// TIA Portal V21 export
// export: Created 2026-11-10T07:35:10.4726746Z, ExportSetting WithDefaults, DisplayName Totally Integrated Automation Portal, DisplayVersion V21 Update 3, DisplayName STEP 7 Professional, DisplayVersion V21 Update 3, DisplayName STEP 7 Safety, DisplayVersion V21, DisplayName Tech WebApplication, DisplayVersion V21, DisplayName WinCC Basic/Comfort/Advanced, DisplayVersion V21 Update 3, DisplayName WinCC Unified, DisplayVersion V21 Update 3
FUNCTION_BLOCK "FB_Lad_ex097"   // FB69, LAD
{ S7_Optimized_Access := 'TRUE' }
VERSION : 0.1
// stored: AutoNumber true, IsIECCheckEnabled false, IsRetainMemResEnabled false, MemoryReserve 100, SetENOAutomatically false, UDAEnableTagReadback false
   VAR_INPUT
      v_req : Bool;
      v_laddr : HW_IO;
      v_recnum : Byte;
      v_ret_val : Int;
   END_VAR
   VAR_OUTPUT
      v_busy : Bool;
   END_VAR
   VAR_IN_OUT
      v_record : Variant;
   END_VAR
BEGIN

REGION Network 1: RD_DPARA - Read module data record asynchronously
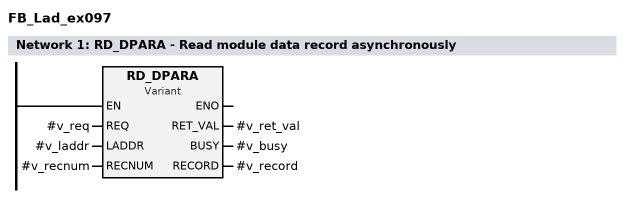
   RUNG wire#powerrail
      { S7_Templates := "[ptr_type := Variant, laddr_type := HW_IO]" } RD_DPARA(REQ := #v_req, LADDR := #v_laddr, RECNUM := #v_recnum, RET_VAL => #v_ret_val, BUSY => #v_busy, RECORD => #v_record)
   END_RUNG
   // the same network as SCL:
   #v_ret_val := RD_DPARA(REQ := #v_req,
                          LADDR := #v_laddr,
                          RECNUM := #v_recnum,
                          BUSY => #v_busy,
                          RECORD => #v_record);
END_REGION
END_FUNCTION_BLOCK
